SUBAPPLICATION Uebung_094b_AX (* Optionsgruppe per VT-Eingabe (Index) auswaehlen: AD_TO_AUI -> AOption_AUI_DEMUX_2 schaltet genau eine von zwei OptionalGroup-SubApps per AOption-Adapter frei (QI anstelle Permit) *)
  (* Standard: 61499-2; Description: Copyright (c) 2026 Meisterschulen am Ostbahnhof This program and the accompanying materials are made available under the terms of the Eclipse Public License 2.0 which is available at https://www.eclipse.org/legal/epl-2.0/ SPDX-License-Identifier: EPL-2.0 *)
  (* Version 1.0, 2026-10-13, Franz Höpfinger, Meisterschulen am Ostbahnhof, initial API and implementation and/or initial documentation *)
  PACKAGE Uebungen;
  IMPORT Uebungen::const::UT::DefaultPool::InputNumber_I1;
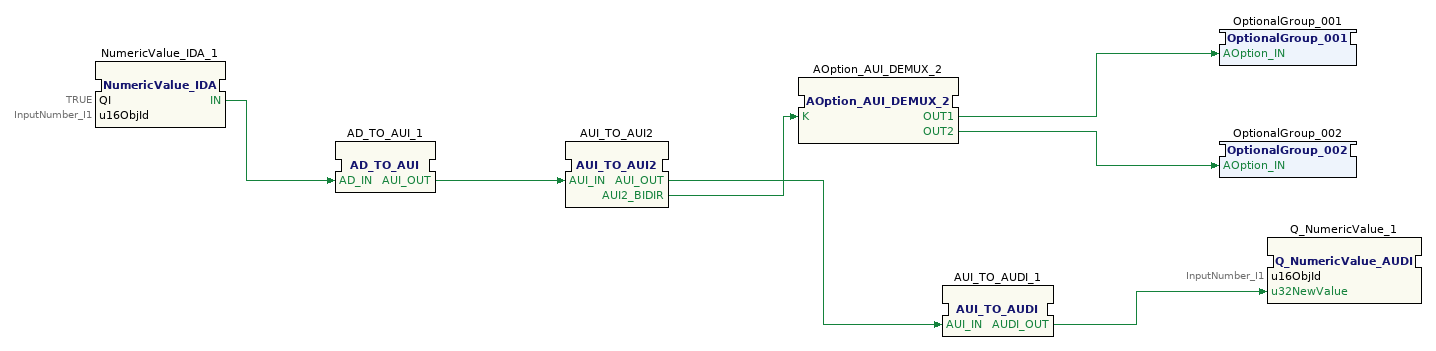
  FBS
    AOption_AUI_DEMUX_2 : Option::selection::AOption_AUI_DEMUX_2;
    Q_NumericValue_1 : isobus::UT::Q::Q_NumericValue_AUDI(u16ObjId := InputNumber_I1);
    AUI_TO_AUDI_1 : adapter::conversion::unidirectional::AUI_TO_AUDI;
    AUI_TO_AUI2 : adapter::conversion::bidirectional::AUI_TO_AUI2;
    AD_TO_AUI_1 : adapter::conversion::unidirectional::AD_TO_AUI;
    NumericValue_IDA_1 : isobus::UT::io::NumericValue::NumericValue_IDA(QI := TRUE, u16ObjId := InputNumber_I1);
  END_FBS
  SUBAPPS
    OptionalGroup_001 : MyLib_AX_Option::sys::OptionalGroup_001;
    OptionalGroup_002 : MyLib_AX_Option::sys::OptionalGroup_002;
  END_SUBAPPS
  ADAPTER_CONNECTIONS
    AOption_AUI_DEMUX_2.OUT1 TO OptionalGroup_001.AOption_IN;
    AOption_AUI_DEMUX_2.OUT2 TO OptionalGroup_002.AOption_IN;
    NumericValue_IDA_1.IN TO AD_TO_AUI_1.AD_IN;
    AD_TO_AUI_1.AUI_OUT TO AUI_TO_AUI2.AUI_IN;
    AUI_TO_AUI2.AUI_OUT TO AUI_TO_AUDI_1.AUI_IN;
    AUI_TO_AUDI_1.AUDI_OUT TO Q_NumericValue_1.u32NewValue;
    AUI_TO_AUI2.AUI2_BIDIR TO AOption_AUI_DEMUX_2.K;
  END_CONNECTIONS
END_SUBAPPLICATION
